FUNCTION_BLOCK ControlPanelOut (* Composite Function Block Type *)
  (* Standard: 61499-2 *)
  (* Version 0.0, 7/2/2026, template *)
  PACKAGE Main;
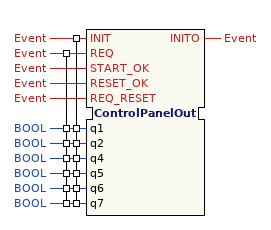
  EVENT_INPUT
    INIT WITH q1, q2, q4, q5, q6, q7; (* Initialization Request *)
    REQ WITH q1, q2, q4, q5, q6, q7; (* Normal Execution Request *)
    START_OK;
    RESET_OK;
    REQ_RESET;
  END_EVENT
  EVENT_OUTPUT
    INITO; (* Initialization Confirm *)
  END_EVENT
  VAR_INPUT
    q1 : BOOL; (* Input event qualifier *)
    q2 : BOOL;
    q4 : BOOL;
    q5 : BOOL;
    q6 : BOOL;
    q7 : BOOL;
  END_VAR
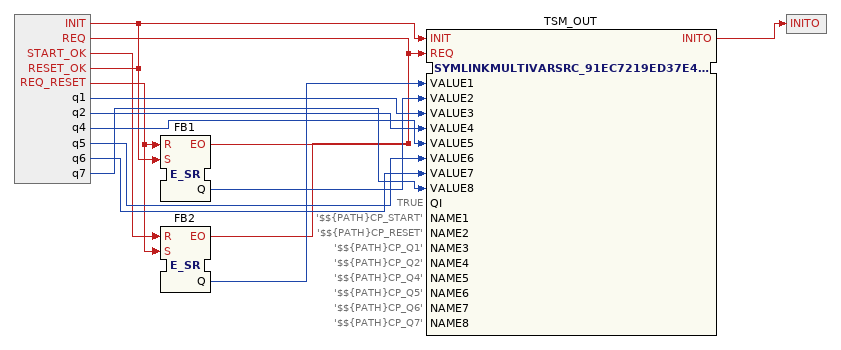
  FBS
    FB1 : E_SR;
    FB2 : E_SR;
    TSM_OUT : SYMLINKMULTIVARSRC_91EC7219ED37E472(QI := TRUE, NAME1 := '$${PATH}CP_START', NAME2 := '$${PATH}CP_RESET', NAME3 := '$${PATH}CP_Q1', NAME4 := '$${PATH}CP_Q2', NAME5 := '$${PATH}CP_Q4', NAME6 := '$${PATH}CP_Q5', NAME7 := '$${PATH}CP_Q6', NAME8 := '$${PATH}CP_Q7'); {SET_ATTRIBUTE(Configuration.GenericFBType.InterfaceParams, Runtime.System#I:=8;VALUE${I$}:BOOL,BOOL,BOOL,BOOL,BOOL,BOOL,BOOL,BOOL)}
  END_FBS
  EVENT_CONNECTIONS
    START_OK TO FB2.R;
    REQ_RESET TO FB1.R;
    REQ_RESET TO FB2.S;
    RESET_OK TO FB1.S;
    INIT TO FB1.S;
    INIT TO TSM_OUT.INIT;
    REQ TO TSM_OUT.REQ;
    FB1.EO TO TSM_OUT.REQ;
    FB2.EO TO TSM_OUT.REQ;
    TSM_OUT.INITO TO INITO;
  END_CONNECTIONS
  DATA_CONNECTIONS
    FB2.Q TO TSM_OUT.VALUE1;
    FB1.Q TO TSM_OUT.VALUE2;
    q1 TO TSM_OUT.VALUE3;
    q2 TO TSM_OUT.VALUE4;
    q4 TO TSM_OUT.VALUE5;
    q5 TO TSM_OUT.VALUE6;
    q6 TO TSM_OUT.VALUE7;
    q7 TO TSM_OUT.VALUE8;
  END_CONNECTIONS
END_FUNCTION_BLOCK
